// TIA Portal V21 export
// export: Created 2026-11-22T04:06:11.2307944Z, ExportSetting WithDefaults, DisplayName Totally Integrated Automation Portal, DisplayVersion V21 Update 3, DisplayName STEP 7 Professional, DisplayVersion V21 Update 3, DisplayName STEP 7 Safety, DisplayVersion V21, DisplayName Tech WebApplication, DisplayVersion V21, DisplayName WinCC Basic/Comfort/Advanced, DisplayVersion V21 Update 3, DisplayName WinCC Unified, DisplayVersion V21 Update 3
ScreenSlidein   NonexNone, Dimension=120, SlideinType=Top, Visibility=FadeOut
  ScreenLayer "Layer_0"
    TextField "SI_Title" at 10,10 size 300x20  StyleItem=Text field, Text="Slide-in screen Top"
    Bar "SI_Bar" at 330,10 size 200x40  CountSubDivisions=5, IntegerDigits=3, LargeTickLabelingStep=1, MaximumValue=5, MinimumValue=-5, Precision=2, StyleItem=Bar
      ProcessValue := D_Pct
    IOField "SI_Value" at 560,10 size 120x30  DataFormat=Decimal, FormatPattern=s99999, Mode=InOutput, StyleItem=I/O field
      ProcessValue := D_Int
